(* IEC 61131-3 sources: plc-st-coding-agent/progress/evidence/f14_v5_public_pilot_20261112/jobs/codex_deepseek-v4pro, 18 files *)

(* ---- public-easy-01.candidate_01.st ---- *)
FUNCTION_BLOCK AutomatedFillingLineControl
VAR_INPUT
    bottleSensor : BOOL;
    cleaningConfirmButton : BOOL;
    fillingConfirmButton : BOOL;
    cappingConfirmButton : BOOL;
    packingConfirmButton : BOOL;
    finishedButton : BOOL;
END_VAR
VAR_OUTPUT
    Pump_Motor : BOOL;
    Filling_Valve : BOOL;
    Capping_Machine : BOOL;
    Packing_Machine : BOOL;
    Completion_Light : BOOL;
END_VAR
VAR
    State : INT := 0;
END_VAR

(* ENGINEERING_CONTRACT
- Pump_Motor: active from bottleSensor detection in Idle and latched through Cleaning; PUB003.
- Pump_Motor: deactivated when cleaningConfirmButton advances to Filling; PUB004.
- Filling_Valve: active from cleaningConfirmButton and held through Filling; PUB004.
- Filling_Valve: deactivated when fillingConfirmButton advances to Capping; PUB005.
- Capping_Machine: active from fillingConfirmButton and held through Capping; PUB005-PUB006.
- Capping_Machine: deactivated when cappingConfirmButton advances to Packing; PUB006.
- Packing_Machine: active from cappingConfirmButton and held through Packing; PUB006-PUB007.
- Packing_Machine: deactivated when packingConfirmButton lights Completion_Light; PUB007.
- Completion_Light: held until finishedButton resets it and returns to Idle; PUB007-PUB008.
- Level-checked inputs; only the current stage consumes its matching confirmation button.
- Same-scan priority: one stage transition per scan; output units are BOOL with no time bounds.
*)

CASE State OF
    0:
        Pump_Motor := FALSE;
        Filling_Valve := FALSE;
        Capping_Machine := FALSE;
        Packing_Machine := FALSE;
        Completion_Light := FALSE;

        IF bottleSensor THEN
            Pump_Motor := TRUE;
            State := 1;
        END_IF;

    1:
        Pump_Motor := TRUE;

        IF cleaningConfirmButton THEN
            Pump_Motor := FALSE;
            Filling_Valve := TRUE;
            State := 2;
        END_IF;

    2:
        Filling_Valve := TRUE;

        IF fillingConfirmButton THEN
            Filling_Valve := FALSE;
            Capping_Machine := TRUE;
            State := 3;
        END_IF;

    3:
        Capping_Machine := TRUE;

        IF cappingConfirmButton THEN
            Capping_Machine := FALSE;
            Packing_Machine := TRUE;
            State := 4;
        END_IF;

    4:
        Packing_Machine := TRUE;

        IF packingConfirmButton THEN
            Packing_Machine := FALSE;
            Completion_Light := TRUE;
            State := 5;
        END_IF;

    5:
        Completion_Light := TRUE;

        IF finishedButton THEN
            Completion_Light := FALSE;
            State := 0;
        END_IF;
END_CASE;

END_FUNCTION_BLOCK

(* ---- public-easy-01.candidate_02.st ---- *)
FUNCTION_BLOCK AutomatedFillingLineControl
VAR_INPUT
    bottleSensor : BOOL;
    cleaningConfirmButton : BOOL;
    fillingConfirmButton : BOOL;
    cappingConfirmButton : BOOL;
    packingConfirmButton : BOOL;
    finishedButton : BOOL;
END_VAR
VAR_OUTPUT
    Pump_Motor : BOOL;
    Filling_Valve : BOOL;
    Capping_Machine : BOOL;
    Packing_Machine : BOOL;
    Completion_Light : BOOL;
END_VAR
VAR
END_VAR

(* ENGINEERING_CONTRACT
- Pump_Motor: activated by bottleSensor, retained/holds until finishedButton reset; PUB003.
- Filling_Valve: activated by cleaningConfirmButton, retained until finishedButton reset; PUB004.
- Capping_Machine: activated by fillingConfirmButton, retained until finishedButton reset; PUB005.
- Packing_Machine: activated by cappingConfirmButton, retained until finishedButton reset; PUB006.
- Completion_Light: activated by packingConfirmButton, retained until finishedButton reset; PUB007.
- finishedButton: explicit common reset for all outputs, applied last in same scan; PUB008.
- Outputs are BOOL; no time bounds. Activation inputs are level-latched, not edge-only.
*)

IF bottleSensor THEN
    Pump_Motor := TRUE;
END_IF;

IF cleaningConfirmButton THEN
    Filling_Valve := TRUE;
END_IF;

IF fillingConfirmButton THEN
    Capping_Machine := TRUE;
END_IF;

IF cappingConfirmButton THEN
    Packing_Machine := TRUE;
END_IF;

IF packingConfirmButton THEN
    Completion_Light := TRUE;
END_IF;

IF finishedButton THEN
    Pump_Motor := FALSE;
    Filling_Valve := FALSE;
    Capping_Machine := FALSE;
    Packing_Machine := FALSE;
    Completion_Light := FALSE;
END_IF;

END_FUNCTION_BLOCK

(* ---- public-easy-01.raw_candidate_01.st ---- *)
FUNCTION_BLOCK AutomatedFillingLineControl
VAR_INPUT
    bottleSensor : BOOL;
    cleaningConfirmButton : BOOL;
    fillingConfirmButton : BOOL;
    cappingConfirmButton : BOOL;
    packingConfirmButton : BOOL;
    finishedButton : BOOL;
END_VAR
VAR_OUTPUT
    Pump_Motor : BOOL;
    Filling_Valve : BOOL;
    Capping_Machine : BOOL;
    Packing_Machine : BOOL;
    Completion_Light : BOOL;
END_VAR
VAR
    State : INT := 0;
END_VAR

(* ENGINEERING_CONTRACT
- Pump_Motor: active from bottleSensor detection in Idle and latched through Cleaning; PUB003.
- Pump_Motor: deactivated when cleaningConfirmButton advances to Filling; PUB004.
- Filling_Valve: active from cleaningConfirmButton and held through Filling; PUB004.
- Filling_Valve: deactivated when fillingConfirmButton advances to Capping; PUB005.
- Capping_Machine: active from fillingConfirmButton and held through Capping; PUB005-PUB006.
- Capping_Machine: deactivated when cappingConfirmButton advances to Packing; PUB006.
- Packing_Machine: active from cappingConfirmButton and held through Packing; PUB006-PUB007.
- Packing_Machine: deactivated when packingConfirmButton lights Completion_Light; PUB007.
- Completion_Light: held until finishedButton resets it and returns to Idle; PUB007-PUB008.
- Level-checked inputs; only the current stage consumes its matching confirmation button.
- Same-scan priority: one stage transition per scan; output units are BOOL with no time bounds.
*)

CASE State OF
    0:
        Pump_Motor := FALSE;
        Filling_Valve := FALSE;
        Capping_Machine := FALSE;
        Packing_Machine := FALSE;
        Completion_Light := FALSE;

        IF bottleSensor THEN
            Pump_Motor := TRUE;
            State := 1;
        END_IF;

    1:
        Pump_Motor := TRUE;

        IF cleaningConfirmButton THEN
            Pump_Motor := FALSE;
            Filling_Valve := TRUE;
            State := 2;
        END_IF;

    2:
        Filling_Valve := TRUE;

        IF fillingConfirmButton THEN
            Filling_Valve := FALSE;
            Capping_Machine := TRUE;
            State := 3;
        END_IF;

    3:
        Capping_Machine := TRUE;

        IF cappingConfirmButton THEN
            Capping_Machine := FALSE;
            Packing_Machine := TRUE;
            State := 4;
        END_IF;

    4:
        Packing_Machine := TRUE;

        IF packingConfirmButton THEN
            Packing_Machine := FALSE;
            Completion_Light := TRUE;
            State := 5;
        END_IF;

    5:
        Completion_Light := TRUE;

        IF finishedButton THEN
            Completion_Light := FALSE;
            State := 0;
        END_IF;
END_CASE;

END_FUNCTION_BLOCK

(* ---- public-easy-01.raw_candidate_02.st ---- *)
FUNCTION_BLOCK AutomatedFillingLineControl
VAR_INPUT
    bottleSensor : BOOL;
    cleaningConfirmButton : BOOL;
    fillingConfirmButton : BOOL;
    cappingConfirmButton : BOOL;
    packingConfirmButton : BOOL;
    finishedButton : BOOL;
END_VAR
VAR_OUTPUT
    Pump_Motor : BOOL;
    Filling_Valve : BOOL;
    Capping_Machine : BOOL;
    Packing_Machine : BOOL;
    Completion_Light : BOOL;
END_VAR
VAR
END_VAR

(* ENGINEERING_CONTRACT
- Pump_Motor: activated by bottleSensor, retained/holds until finishedButton reset; PUB003.
- Filling_Valve: activated by cleaningConfirmButton, retained until finishedButton reset; PUB004.
- Capping_Machine: activated by fillingConfirmButton, retained until finishedButton reset; PUB005.
- Packing_Machine: activated by cappingConfirmButton, retained until finishedButton reset; PUB006.
- Completion_Light: activated by packingConfirmButton, retained until finishedButton reset; PUB007.
- finishedButton: explicit common reset for all outputs, applied last in same scan; PUB008.
- Outputs are BOOL; no time bounds. Activation inputs are level-latched, not edge-only.
*)

IF bottleSensor THEN
    Pump_Motor := TRUE;
END_IF;

IF cleaningConfirmButton THEN
    Filling_Valve := TRUE;
END_IF;

IF fillingConfirmButton THEN
    Capping_Machine := TRUE;
END_IF;

IF cappingConfirmButton THEN
    Packing_Machine := TRUE;
END_IF;

IF packingConfirmButton THEN
    Completion_Light := TRUE;
END_IF;

IF finishedButton THEN
    Pump_Motor := FALSE;
    Filling_Valve := FALSE;
    Capping_Machine := FALSE;
    Packing_Machine := FALSE;
    Completion_Light := FALSE;
END_IF;

END_FUNCTION_BLOCK

(* ---- public-easy-04.candidate_01.st ---- *)
(*
ENGINEERING_CONTRACT
VFD_RUN [PUB002,PUB003,PUB006]: TRUE only while PASTE_E_STOP_NC=TRUE and the viscosity debounce timer has elapsed; same-scan emergency stop drops the run command and clears incomplete debounce timing; power-up state is OFF.
Debounce [PUB002,PUB003]: timer IN uses VISCOSITY_OK AND PASTE_E_STOP_NC with PT=DebounceTime; a FALSE viscosity input invalidates immediately, and a FALSE emergency stop resets incomplete timing.
Runtime [PUB004,PUB006]: adds TIME_TO_LTIME(CycleTime) once per invocation only while VFD_RUN=TRUE; preserves the accumulated value while stopped; starts at 0 ns.
Maintenance [PUB005,PUB006]: PUMP_MAINT_DUE becomes TRUE when accumulated runtime reaches 500 h; it is informational only, remains TRUE because runtime is monotonic, and does not affect run or safety logic; starts FALSE.
Units/boundaries: maintenance threshold uses T#500h with >= comparison; CycleTime and DebounceTime are assumed positive.
Unspecified: no reset is defined for accumulated runtime or the maintenance indication; non-positive input times follow normal TON/add behavior without additional clamping.
*)
FUNCTION_BLOCK JamPumpControl
VAR_INPUT
    VISCOSITY_OK : BOOL;
    PASTE_E_STOP_NC : BOOL;
    DebounceTime : TIME;
    CycleTime : TIME;
END_VAR
VAR_OUTPUT
    VFD_RUN : BOOL;
    PUMP_MAINT_DUE : BOOL;
    PUMP_RUNTIME_ACC : LTIME;
END_VAR
VAR
    tonViscosity : TON;
    RuntimeAcc : LTIME := LTIME#0s;
    MAINT_THRESHOLD : TIME := T#500h;
END_VAR

tonViscosity(IN := (VISCOSITY_OK AND PASTE_E_STOP_NC), PT := DebounceTime);

VFD_RUN := PASTE_E_STOP_NC AND tonViscosity.Q;

IF VFD_RUN THEN
    RuntimeAcc := RuntimeAcc + TIME_TO_LTIME(CycleTime);
END_IF;

PUMP_RUNTIME_ACC := RuntimeAcc;
PUMP_MAINT_DUE := PUMP_RUNTIME_ACC >= TIME_TO_LTIME(MAINT_THRESHOLD);

END_FUNCTION_BLOCK

(* ---- public-easy-04.raw_candidate_01.st ---- *)
(*
ENGINEERING_CONTRACT
VFD_RUN [PUB002,PUB003,PUB006]: TRUE only while PASTE_E_STOP_NC=TRUE and the viscosity debounce timer has elapsed; same-scan emergency stop drops the run command and clears incomplete debounce timing; power-up state is OFF.
Debounce [PUB002,PUB003]: timer IN uses VISCOSITY_OK AND PASTE_E_STOP_NC with PT=DebounceTime; a FALSE viscosity input invalidates immediately, and a FALSE emergency stop resets incomplete timing.
Runtime [PUB004,PUB006]: adds TIME_TO_LTIME(CycleTime) once per invocation only while VFD_RUN=TRUE; preserves the accumulated value while stopped; starts at 0 ns.
Maintenance [PUB005,PUB006]: PUMP_MAINT_DUE becomes TRUE when accumulated runtime reaches 500 h; it is informational only, remains TRUE because runtime is monotonic, and does not affect run or safety logic; starts FALSE.
Units/boundaries: maintenance threshold uses T#500h with >= comparison; CycleTime and DebounceTime are assumed positive.
Unspecified: no reset is defined for accumulated runtime or the maintenance indication; non-positive input times follow normal TON/add behavior without additional clamping.
*)
FUNCTION_BLOCK JamPumpControl
VAR_INPUT
    VISCOSITY_OK : BOOL;
    PASTE_E_STOP_NC : BOOL;
    DebounceTime : TIME;
    CycleTime : TIME;
END_VAR
VAR_OUTPUT
    VFD_RUN : BOOL;
    PUMP_MAINT_DUE : BOOL;
    PUMP_RUNTIME_ACC : LTIME;
END_VAR
VAR
    tonViscosity : TON;
    RuntimeAcc : LTIME := LTIME#0s;
    MAINT_THRESHOLD : TIME := T#500h;
END_VAR

tonViscosity(IN := (VISCOSITY_OK AND PASTE_E_STOP_NC), PT := DebounceTime);

VFD_RUN := PASTE_E_STOP_NC AND tonViscosity.Q;

IF VFD_RUN THEN
    RuntimeAcc := RuntimeAcc + TIME_TO_LTIME(CycleTime);
END_IF;

PUMP_RUNTIME_ACC := RuntimeAcc;
PUMP_MAINT_DUE := PUMP_RUNTIME_ACC >= TIME_TO_LTIME(MAINT_THRESHOLD);

END_FUNCTION_BLOCK

(* ---- public-hard-03.candidate_01.st ---- *)
TYPE ST_Recipe :
STRUCT
    recipeID : INT;
    ingredientType : INT;
    ingredientRatio : REAL;
    productionTemperature : REAL;
END_STRUCT
END_TYPE;

FUNCTION_BLOCK RecipeManagementSystem
(*
ENGINEERING_CONTRACT
- Operations are level-triggered; no edge or latch storage is added (PUB002-PUB006).
- recipeAdded/Deleted/Modified are active only during a successful selected scan; otherwise cleared.
- error/status clear each scan unless the selected operation reports a failure.
- Query retains the last successful recipeQueryResult; a missing recipe leaves it unchanged (PUB009).
- Add checks duplicate first, then smallest empty index, otherwise 16#8002/16#8003 (PUB010).
- Delete clears only recipeID in the matched slot (PUB011).
- Modify replaces the whole matched ST_Recipe with recipeIn (PUB012).
- recipeID=0 denotes an empty slot; searches ignore such slots (PUB008).
- Simultaneous requests use priority add > delete > modify > query (unspecified by task).
*)
VAR_INPUT
    addRecipe : BOOL;
    deleteRecipe : BOOL;
    modifyRecipe : BOOL;
    queryRecipe : BOOL;
    recipeIn : ST_Recipe;
END_VAR
VAR_OUTPUT
    recipeAdded : BOOL;
    recipeDeleted : BOOL;
    recipeModified : BOOL;
    recipeQueryResult : ST_Recipe;
    error : BOOL;
    status : WORD;
END_VAR
VAR_IN_OUT
    recipe : ARRAY[1..10] OF ST_Recipe;
END_VAR
VAR
    i : INT;
    foundIndex : INT;
    emptyIndex : INT;
    found : BOOL;
    emptyFound : BOOL;
END_VAR

recipeAdded := FALSE;
recipeDeleted := FALSE;
recipeModified := FALSE;
error := FALSE;
status := 0;

IF addRecipe THEN
    found := FALSE;
    foundIndex := 0;
    FOR i := 1 TO 10 DO
        IF (recipe[i].recipeID <> 0) AND (recipe[i].recipeID = recipeIn.recipeID) THEN
            found := TRUE;
            foundIndex := i;
            EXIT;
        END_IF;
    END_FOR;

    IF found THEN
        error := TRUE;
        status := WORD#16#8002;
    ELSE
        emptyFound := FALSE;
        emptyIndex := 0;
        FOR i := 1 TO 10 DO
            IF recipe[i].recipeID = 0 THEN
                emptyFound := TRUE;
                emptyIndex := i;
                EXIT;
            END_IF;
        END_FOR;

        IF NOT emptyFound THEN
            error := TRUE;
            status := WORD#16#8003;
        ELSE
            recipe[emptyIndex].recipeID := recipeIn.recipeID;
            recipe[emptyIndex].ingredientType := recipeIn.ingredientType;
            recipe[emptyIndex].ingredientRatio := recipeIn.ingredientRatio;
            recipe[emptyIndex].productionTemperature := recipeIn.productionTemperature;
            recipeAdded := TRUE;
            error := FALSE;
            status := 0;
        END_IF;
    END_IF;

ELSIF deleteRecipe THEN
    found := FALSE;
    foundIndex := 0;
    FOR i := 1 TO 10 DO
        IF (recipe[i].recipeID <> 0) AND (recipe[i].recipeID = recipeIn.recipeID) THEN
            found := TRUE;
            foundIndex := i;
            EXIT;
        END_IF;
    END_FOR;

    IF NOT found THEN
        error := TRUE;
        status := WORD#16#8004;
    ELSE
        recipe[foundIndex].recipeID := 0;
        recipeDeleted := TRUE;
        error := FALSE;
        status := 0;
    END_IF;

ELSIF modifyRecipe THEN
    found := FALSE;
    foundIndex := 0;
    FOR i := 1 TO 10 DO
        IF (recipe[i].recipeID <> 0) AND (recipe[i].recipeID = recipeIn.recipeID) THEN
            found := TRUE;
            foundIndex := i;
            EXIT;
        END_IF;
    END_FOR;

    IF NOT found THEN
        error := TRUE;
        status := WORD#16#8005;
    ELSE
        recipe[foundIndex] := recipeIn;
        recipeModified := TRUE;
        error := FALSE;
        status := 0;
    END_IF;

ELSIF queryRecipe THEN
    found := FALSE;
    foundIndex := 0;
    FOR i := 1 TO 10 DO
        IF (recipe[i].recipeID <> 0) AND (recipe[i].recipeID = recipeIn.recipeID) THEN
            found := TRUE;
            foundIndex := i;
            EXIT;
        END_IF;
    END_FOR;

    IF NOT found THEN
        error := TRUE;
        status := WORD#16#8001;
    ELSE
        recipeQueryResult := recipe[foundIndex];
        error := FALSE;
        status := 0;
    END_IF;
END_IF;

END_FUNCTION_BLOCK

(* ---- public-hard-03.candidate_02.st ---- *)
TYPE ST_Recipe :
STRUCT
    recipeID : INT;
    ingredientType : INT;
    ingredientRatio : REAL;
    productionTemperature : REAL;
END_STRUCT
END_TYPE;

FUNCTION_BLOCK RecipeManagementSystem
(*
ENGINEERING_CONTRACT
- Request inputs are level-triggered; no edge or latch storage is added.
- recipeAdded/recipeDeleted/recipeModified are true only on a successful scan of the matching request, otherwise false.
- error/status clear at scan start; any failed request in the scan sets them.
- Query success overwrites recipeQueryResult; a failed query leaves it unchanged.
- Add checks duplicate first, then finds the smallest empty index, then checks full database.
- Delete clears only recipeID in the matched slot.
- Modify replaces the entire matched ST_Recipe with recipeIn.
- Empty slots are identified by recipeID = 0 and are ignored during normal searches.
- Simultaneous requests are unspecified; they are evaluated in interface order add/delete/modify/query.
*)
VAR_INPUT
    addRecipe : BOOL;
    deleteRecipe : BOOL;
    modifyRecipe : BOOL;
    queryRecipe : BOOL;
    recipeIn : ST_Recipe;
END_VAR
VAR_OUTPUT
    recipeAdded : BOOL;
    recipeDeleted : BOOL;
    recipeModified : BOOL;
    recipeQueryResult : ST_Recipe;
    error : BOOL;
    status : WORD;
END_VAR
VAR_IN_OUT
    recipe : ARRAY[1..10] OF ST_Recipe;
END_VAR
VAR
    i : INT;
    foundIndex : INT;
    emptyIndex : INT;
    found : BOOL;
    emptyFound : BOOL;
END_VAR

recipeAdded := FALSE;
recipeDeleted := FALSE;
recipeModified := FALSE;
error := FALSE;
status := 0;

IF addRecipe THEN
    found := FALSE;
    foundIndex := 0;
    FOR i := 1 TO 10 DO
        IF (recipe[i].recipeID <> 0) AND (recipe[i].recipeID = recipeIn.recipeID) THEN
            found := TRUE;
            foundIndex := i;
            EXIT;
        END_IF;
    END_FOR;

    IF found THEN
        error := TRUE;
        status := WORD#16#8002;
    ELSE
        emptyFound := FALSE;
        emptyIndex := 0;
        FOR i := 1 TO 10 DO
            IF recipe[i].recipeID = 0 THEN
                emptyFound := TRUE;
                emptyIndex := i;
                EXIT;
            END_IF;
        END_FOR;

        IF NOT emptyFound THEN
            error := TRUE;
            status := WORD#16#8003;
        ELSE
            recipe[emptyIndex].recipeID := recipeIn.recipeID;
            recipe[emptyIndex].ingredientType := recipeIn.ingredientType;
            recipe[emptyIndex].ingredientRatio := recipeIn.ingredientRatio;
            recipe[emptyIndex].productionTemperature := recipeIn.productionTemperature;
            recipeAdded := TRUE;
        END_IF;
    END_IF;
END_IF;

IF deleteRecipe THEN
    found := FALSE;
    foundIndex := 0;
    FOR i := 1 TO 10 DO
        IF (recipe[i].recipeID <> 0) AND (recipe[i].recipeID = recipeIn.recipeID) THEN
            found := TRUE;
            foundIndex := i;
            EXIT;
        END_IF;
    END_FOR;

    IF NOT found THEN
        error := TRUE;
        status := WORD#16#8004;
    ELSE
        recipe[foundIndex].recipeID := 0;
        recipeDeleted := TRUE;
    END_IF;
END_IF;

IF modifyRecipe THEN
    found := FALSE;
    foundIndex := 0;
    FOR i := 1 TO 10 DO
        IF (recipe[i].recipeID <> 0) AND (recipe[i].recipeID = recipeIn.recipeID) THEN
            found := TRUE;
            foundIndex := i;
            EXIT;
        END_IF;
    END_FOR;

    IF NOT found THEN
        error := TRUE;
        status := WORD#16#8005;
    ELSE
        recipe[foundIndex] := recipeIn;
        recipeModified := TRUE;
    END_IF;
END_IF;

IF queryRecipe THEN
    found := FALSE;
    foundIndex := 0;
    FOR i := 1 TO 10 DO
        IF (recipe[i].recipeID <> 0) AND (recipe[i].recipeID = recipeIn.recipeID) THEN
            found := TRUE;
            foundIndex := i;
            EXIT;
        END_IF;
    END_FOR;

    IF NOT found THEN
        error := TRUE;
        status := WORD#16#8001;
    ELSE
        recipeQueryResult := recipe[foundIndex];
    END_IF;
END_IF;

END_FUNCTION_BLOCK

(* ---- public-hard-03.raw_candidate_01.st ---- *)
TYPE ST_Recipe :
STRUCT
    recipeID : INT;
    ingredientType : INT;
    ingredientRatio : REAL;
    productionTemperature : REAL;
END_STRUCT
END_TYPE

FUNCTION_BLOCK RecipeManagementSystem
(*
ENGINEERING_CONTRACT
- Operations are level-triggered; no edge or latch storage is added (PUB002-PUB006).
- recipeAdded/Deleted/Modified are active only during a successful selected scan; otherwise cleared.
- error/status clear each scan unless the selected operation reports a failure.
- Query retains the last successful recipeQueryResult; a missing recipe leaves it unchanged (PUB009).
- Add checks duplicate first, then smallest empty index, otherwise 16#8002/16#8003 (PUB010).
- Delete clears only recipeID in the matched slot (PUB011).
- Modify replaces the whole matched ST_Recipe with recipeIn (PUB012).
- recipeID=0 denotes an empty slot; searches ignore such slots (PUB008).
- Simultaneous requests use priority add > delete > modify > query (unspecified by task).
*)
VAR_INPUT
    addRecipe : BOOL;
    deleteRecipe : BOOL;
    modifyRecipe : BOOL;
    queryRecipe : BOOL;
    recipeIn : ST_Recipe;
END_VAR
VAR_OUTPUT
    recipeAdded : BOOL;
    recipeDeleted : BOOL;
    recipeModified : BOOL;
    recipeQueryResult : ST_Recipe;
    error : BOOL;
    status : WORD;
END_VAR
VAR_IN_OUT
    recipe : ARRAY[1..10] OF ST_Recipe;
END_VAR
VAR
    i : INT;
    foundIndex : INT;
    emptyIndex : INT;
    found : BOOL;
    emptyFound : BOOL;
END_VAR

recipeAdded := FALSE;
recipeDeleted := FALSE;
recipeModified := FALSE;
error := FALSE;
status := 0;

IF addRecipe THEN
    found := FALSE;
    foundIndex := 0;
    FOR i := 1 TO 10 DO
        IF (recipe[i].recipeID <> 0) AND (recipe[i].recipeID = recipeIn.recipeID) THEN
            found := TRUE;
            foundIndex := i;
            EXIT;
        END_IF;
    END_FOR;

    IF found THEN
        error := TRUE;
        status := WORD#16#8002;
    ELSE
        emptyFound := FALSE;
        emptyIndex := 0;
        FOR i := 1 TO 10 DO
            IF recipe[i].recipeID = 0 THEN
                emptyFound := TRUE;
                emptyIndex := i;
                EXIT;
            END_IF;
        END_FOR;

        IF NOT emptyFound THEN
            error := TRUE;
            status := WORD#16#8003;
        ELSE
            recipe[emptyIndex].recipeID := recipeIn.recipeID;
            recipe[emptyIndex].ingredientType := recipeIn.ingredientType;
            recipe[emptyIndex].ingredientRatio := recipeIn.ingredientRatio;
            recipe[emptyIndex].productionTemperature := recipeIn.productionTemperature;
            recipeAdded := TRUE;
            error := FALSE;
            status := 0;
        END_IF;
    END_IF;

ELSIF deleteRecipe THEN
    found := FALSE;
    foundIndex := 0;
    FOR i := 1 TO 10 DO
        IF (recipe[i].recipeID <> 0) AND (recipe[i].recipeID = recipeIn.recipeID) THEN
            found := TRUE;
            foundIndex := i;
            EXIT;
        END_IF;
    END_FOR;

    IF NOT found THEN
        error := TRUE;
        status := WORD#16#8004;
    ELSE
        recipe[foundIndex].recipeID := 0;
        recipeDeleted := TRUE;
        error := FALSE;
        status := 0;
    END_IF;

ELSIF modifyRecipe THEN
    found := FALSE;
    foundIndex := 0;
    FOR i := 1 TO 10 DO
        IF (recipe[i].recipeID <> 0) AND (recipe[i].recipeID = recipeIn.recipeID) THEN
            found := TRUE;
            foundIndex := i;
            EXIT;
        END_IF;
    END_FOR;

    IF NOT found THEN
        error := TRUE;
        status := WORD#16#8005;
    ELSE
        recipe[foundIndex] := recipeIn;
        recipeModified := TRUE;
        error := FALSE;
        status := 0;
    END_IF;

ELSIF queryRecipe THEN
    found := FALSE;
    foundIndex := 0;
    FOR i := 1 TO 10 DO
        IF (recipe[i].recipeID <> 0) AND (recipe[i].recipeID = recipeIn.recipeID) THEN
            found := TRUE;
            foundIndex := i;
            EXIT;
        END_IF;
    END_FOR;

    IF NOT found THEN
        error := TRUE;
        status := WORD#16#8001;
    ELSE
        recipeQueryResult := recipe[foundIndex];
        error := FALSE;
        status := 0;
    END_IF;
END_IF;

END_FUNCTION_BLOCK

(* ---- public-hard-03.raw_candidate_02.st ---- *)
TYPE ST_Recipe :
STRUCT
    recipeID : INT;
    ingredientType : INT;
    ingredientRatio : REAL;
    productionTemperature : REAL;
END_STRUCT
END_TYPE;

FUNCTION_BLOCK RecipeManagementSystem
(*
ENGINEERING_CONTRACT
- Request inputs are level-triggered; no edge or latch storage is added.
- recipeAdded/recipeDeleted/recipeModified are true only on a successful scan of the matching request, otherwise false.
- error/status clear at scan start; any failed request in the scan sets them.
- Query success overwrites recipeQueryResult; a failed query leaves it unchanged.
- Add checks duplicate first, then finds the smallest empty index, then checks full database.
- Delete clears only recipeID in the matched slot.
- Modify replaces the entire matched ST_Recipe with recipeIn.
- Empty slots are identified by recipeID = 0 and are ignored during normal searches.
- Simultaneous requests are unspecified; they are evaluated in interface order add/delete/modify/query.
*)
VAR_INPUT
    addRecipe : BOOL;
    deleteRecipe : BOOL;
    modifyRecipe : BOOL;
    queryRecipe : BOOL;
    recipeIn : ST_Recipe;
END_VAR
VAR_OUTPUT
    recipeAdded : BOOL;
    recipeDeleted : BOOL;
    recipeModified : BOOL;
    recipeQueryResult : ST_Recipe;
    error : BOOL;
    status : WORD;
END_VAR
VAR_IN_OUT
    recipe : ARRAY[1..10] OF ST_Recipe;
END_VAR
VAR
    i : INT;
    foundIndex : INT;
    emptyIndex : INT;
    found : BOOL;
    emptyFound : BOOL;
END_VAR

recipeAdded := FALSE;
recipeDeleted := FALSE;
recipeModified := FALSE;
error := FALSE;
status := 0;

IF addRecipe THEN
    found := FALSE;
    foundIndex := 0;
    FOR i := 1 TO 10 DO
        IF (recipe[i].recipeID <> 0) AND (recipe[i].recipeID = recipeIn.recipeID) THEN
            found := TRUE;
            foundIndex := i;
            EXIT;
        END_IF;
    END_FOR;

    IF found THEN
        error := TRUE;
        status := WORD#16#8002;
    ELSE
        emptyFound := FALSE;
        emptyIndex := 0;
        FOR i := 1 TO 10 DO
            IF recipe[i].recipeID = 0 THEN
                emptyFound := TRUE;
                emptyIndex := i;
                EXIT;
            END_IF;
        END_FOR;

        IF NOT emptyFound THEN
            error := TRUE;
            status := WORD#16#8003;
        ELSE
            recipe[emptyIndex].recipeID := recipeIn.recipeID;
            recipe[emptyIndex].ingredientType := recipeIn.ingredientType;
            recipe[emptyIndex].ingredientRatio := recipeIn.ingredientRatio;
            recipe[emptyIndex].productionTemperature := recipeIn.productionTemperature;
            recipeAdded := TRUE;
        END_IF;
    END_IF;
END_IF;

IF deleteRecipe THEN
    found := FALSE;
    foundIndex := 0;
    FOR i := 1 TO 10 DO
        IF (recipe[i].recipeID <> 0) AND (recipe[i].recipeID = recipeIn.recipeID) THEN
            found := TRUE;
            foundIndex := i;
            EXIT;
        END_IF;
    END_FOR;

    IF NOT found THEN
        error := TRUE;
        status := WORD#16#8004;
    ELSE
        recipe[foundIndex].recipeID := 0;
        recipeDeleted := TRUE;
    END_IF;
END_IF;

IF modifyRecipe THEN
    found := FALSE;
    foundIndex := 0;
    FOR i := 1 TO 10 DO
        IF (recipe[i].recipeID <> 0) AND (recipe[i].recipeID = recipeIn.recipeID) THEN
            found := TRUE;
            foundIndex := i;
            EXIT;
        END_IF;
    END_FOR;

    IF NOT found THEN
        error := TRUE;
        status := WORD#16#8005;
    ELSE
        recipe[foundIndex] := recipeIn;
        recipeModified := TRUE;
    END_IF;
END_IF;

IF queryRecipe THEN
    found := FALSE;
    foundIndex := 0;
    FOR i := 1 TO 10 DO
        IF (recipe[i].recipeID <> 0) AND (recipe[i].recipeID = recipeIn.recipeID) THEN
            found := TRUE;
            foundIndex := i;
            EXIT;
        END_IF;
    END_FOR;

    IF NOT found THEN
        error := TRUE;
        status := WORD#16#8001;
    ELSE
        recipeQueryResult := recipe[foundIndex];
    END_IF;
END_IF;

END_FUNCTION_BLOCK

(* ---- public-medium-03.candidate_01.st ---- *)
(* ENGINEERING_CONTRACT
   average: recomputed each scan for active stored samples; 0.0 when no samples or after reset. Units follow value.
   windowSizeReached: TRUE iff stored valid sample count >= current valid windowSize; cleared by reset and on invalid window.
   error/status: enabled by windowSize outside 1..100; status 16#8200, otherwise 16#0000 (PUB004/PUB006/PUB007).
   same-scan priority: level-true reset first, then window validation, then cyclic or rising-edge sample; cyclic TRUE ignores trigger edge (PUB002/PUB003).
   reset: explicit level-true clear of stored samples, count, average, and reached state; no same-scan sample after reset.
   trigger: internal rising-edge detector; each valid, non-reset rising edge adds one value.
   retention: valid stored samples persist without reset; dynamic window resizing uses the newest min(validCount, windowSize) samples.
   boundaries: windowSize [1,100], storage capacity 100; average is LREAL mean with no unit conversion.
*)
FUNCTION_BLOCK FB
VAR_INPUT
    cyclicExecution : BOOL;
    trigger : BOOL;
    value : LREAL;
    windowSize : INT;
    reset : BOOL;
END_VAR
VAR_OUTPUT
    average : LREAL;
    windowSizeReached : BOOL;
    error : BOOL;
    status : WORD;
END_VAR
VAR
    buffer : ARRAY[0..99] OF LREAL;
    nextIndex : INT := 0;
    validCount : INT := 0;
    triggerPrevious : BOOL;
    triggerRising : BOOL;
    activeWindow : INT;
    startIndex : INT;
    loopIndex : INT;
    sumValue : LREAL;
END_VAR

triggerRising := trigger AND NOT triggerPrevious;
triggerPrevious := trigger;

IF reset THEN
    validCount := 0;
    nextIndex := 0;
    average := 0.0;
    windowSizeReached := FALSE;
END_IF;

IF (windowSize < 1) OR (windowSize > 100) THEN
    error := TRUE;
    status := 16#8200;
    average := 0.0;
    windowSizeReached := FALSE;
ELSE
    error := FALSE;
    status := 16#0000;

    IF NOT reset THEN
        IF cyclicExecution OR triggerRising THEN
            buffer[nextIndex] := value;
            nextIndex := nextIndex + 1;

            IF nextIndex > 99 THEN
                nextIndex := 0;
            END_IF;

            IF validCount < 100 THEN
                validCount := validCount + 1;
            END_IF;
        END_IF;
    END_IF;

    activeWindow := windowSize;
    IF activeWindow > validCount THEN
        activeWindow := validCount;
    END_IF;

    IF activeWindow > 0 THEN
        sumValue := 0.0;
        FOR loopIndex := 0 TO activeWindow - 1 DO
            startIndex := nextIndex - 1 - loopIndex;
            IF startIndex < 0 THEN
                startIndex := startIndex + 100;
            END_IF;
            sumValue := sumValue + buffer[startIndex];
        END_FOR;
        average := sumValue / INT_TO_LREAL(activeWindow);
    ELSE
        average := 0.0;
    END_IF;

    windowSizeReached := validCount >= windowSize;
END_IF;
END_FUNCTION_BLOCK

(* ---- public-medium-03.raw_candidate_01.st ---- *)
(* ENGINEERING_CONTRACT
   average: recomputed each scan for active stored samples; 0.0 when no samples or after reset. Units follow value.
   windowSizeReached: TRUE iff stored valid sample count >= current valid windowSize; cleared by reset and on invalid window.
   error/status: enabled by windowSize outside 1..100; status 16#8200, otherwise 16#0000 (PUB004/PUB006/PUB007).
   same-scan priority: level-true reset first, then window validation, then cyclic or rising-edge sample; cyclic TRUE ignores trigger edge (PUB002/PUB003).
   reset: explicit level-true clear of stored samples, count, average, and reached state; no same-scan sample after reset.
   trigger: internal rising-edge detector; each valid, non-reset rising edge adds one value.
   retention: valid stored samples persist without reset; dynamic window resizing uses the newest min(validCount, windowSize) samples.
   boundaries: windowSize [1,100], storage capacity 100; average is LREAL mean with no unit conversion.
*)
FUNCTION_BLOCK FB
VAR_INPUT
    cyclicExecution : BOOL;
    trigger : BOOL;
    value : LREAL;
    windowSize : INT;
    reset : BOOL;
END_VAR
VAR_OUTPUT
    average : LREAL;
    windowSizeReached : BOOL;
    error : BOOL;
    status : WORD;
END_VAR
VAR
    buffer : ARRAY[0..99] OF LREAL;
    nextIndex : INT := 0;
    validCount : INT := 0;
    triggerPrevious : BOOL;
    triggerRising : BOOL;
    activeWindow : INT;
    startIndex : INT;
    loopIndex : INT;
    sumValue : LREAL;
END_VAR

triggerRising := trigger AND NOT triggerPrevious;
triggerPrevious := trigger;

IF reset THEN
    validCount := 0;
    nextIndex := 0;
    average := 0.0;
    windowSizeReached := FALSE;
END_IF;

IF (windowSize < 1) OR (windowSize > 100) THEN
    error := TRUE;
    status := 16#8200;
    average := 0.0;
    windowSizeReached := FALSE;
ELSE
    error := FALSE;
    status := 16#0000;

    IF NOT reset THEN
        IF cyclicExecution OR triggerRising THEN
            buffer[nextIndex] := value;
            nextIndex := nextIndex + 1;

            IF nextIndex > 99 THEN
                nextIndex := 0;
            END_IF;

            IF validCount < 100 THEN
                validCount := validCount + 1;
            END_IF;
        END_IF;
    END_IF;

    activeWindow := windowSize;
    IF activeWindow > validCount THEN
        activeWindow := validCount;
    END_IF;

    IF activeWindow > 0 THEN
        sumValue := 0.0;
        FOR loopIndex := 0 TO activeWindow - 1 DO
            startIndex := nextIndex - 1 - loopIndex;
            IF startIndex < 0 THEN
                startIndex := startIndex + 100;
            END_IF;
            sumValue := sumValue + buffer[startIndex];
        END_FOR;
        average := sumValue / INT_TO_LREAL(activeWindow);
    ELSE
        average := 0.0;
    END_IF;

    windowSizeReached := validCount >= windowSize;
END_IF;
END_FUNCTION_BLOCK

(* ---- public-medium-04.candidate_01.st ---- *)
FUNCTION_BLOCK FB_TemperatureControl
VAR_INPUT
    TemperatureSensorInput : REAL;
    SetTemperature : REAL;
END_VAR
VAR_OUTPUT
    CurrentTemperature : REAL;
    SetTempDisplay : REAL;
    HeaterStatus : BOOL;
    OverheatProtection : BOOL;
    HeaterOutput : BOOL;
END_VAR
VAR
    SensorFault : BOOL;
    HeatRunTimer : TON;
    CoolDownTimer : TON;
END_VAR

(* ENGINEERING_CONTRACT
- CurrentTemperature/SetTempDisplay: copied from inputs every scan (PUB001, PUB002, PUB007); no retention; REAL.
- HeaterStatus: ON only while HeaterOutput is ON; no latch; cleared with heater OFF, overheat, or fault; same-scan as HeaterOutput; BOOL.
- OverheatProtection: latched when continuous heater run reaches >= T#5S (PUB006); held during T#3S cooldown; auto-clears after cooldown; BOOL.
- HeaterOutput: ON when no fault and actual < set (PUB003, PUB004); OFF when actual >= set, sensor fault, or protection (PUB005, PUB007, PUB008).
- SensorFault: TRUE when input < 0.0 or > 100.0 (PUB008); forces heater OFF; does not reset an active overheat cooldown.
- Unspecified: actual = set is interpreted as OFF; no hysteresis; after T#3S cooldown, normal control resumes automatically.
*)

CurrentTemperature := TemperatureSensorInput;
SetTempDisplay := SetTemperature;

SensorFault := (TemperatureSensorInput < 0.0) OR (TemperatureSensorInput > 100.0);

IF SensorFault THEN
    HeaterOutput := FALSE;
    HeaterStatus := FALSE;
    HeatRunTimer(IN := FALSE, PT := T#5S);

    IF OverheatProtection THEN
        CoolDownTimer(IN := TRUE, PT := T#3S);
        IF CoolDownTimer.Q THEN
            OverheatProtection := FALSE;
        END_IF;
    ELSE
        CoolDownTimer(IN := FALSE, PT := T#3S);
    END_IF;

ELSE
    IF OverheatProtection THEN
        HeaterOutput := FALSE;
        HeaterStatus := FALSE;
        HeatRunTimer(IN := FALSE, PT := T#5S);
        CoolDownTimer(IN := TRUE, PT := T#3S);

        IF CoolDownTimer.Q THEN
            OverheatProtection := FALSE;
        END_IF;

    ELSE
        IF TemperatureSensorInput < SetTemperature THEN
            HeaterOutput := TRUE;
            HeaterStatus := TRUE;
            HeatRunTimer(IN := TRUE, PT := T#5S);
            CoolDownTimer(IN := FALSE, PT := T#3S);

            IF HeatRunTimer.Q THEN
                OverheatProtection := TRUE;
                HeaterOutput := FALSE;
                HeaterStatus := FALSE;
            END_IF;

        ELSE
            HeaterOutput := FALSE;
            HeaterStatus := FALSE;
            HeatRunTimer(IN := FALSE, PT := T#5S);
            CoolDownTimer(IN := FALSE, PT := T#3S);
        END_IF;
    END_IF;
END_IF;

END_FUNCTION_BLOCK

(* ---- public-medium-04.candidate_02.st ---- *)
FUNCTION_BLOCK FB_TemperatureControl
VAR_INPUT
    TemperatureSensorInput : REAL;
    SetTemperature : REAL;
END_VAR
VAR_OUTPUT
    CurrentTemperature : REAL;
    SetTempDisplay : REAL;
    HeaterStatus : BOOL;
    OverheatProtection : BOOL;
    HeaterOutput : BOOL;
END_VAR
VAR
    SensorFault : BOOL;
    FreeClock : TON;
    HeatStartTime : TIME;
    HeatWasRunning : BOOL;
    HeatElapsed : TIME;
    CooldownStartTime : TIME;
    CoolElapsed : TIME;
END_VAR

(* ENGINEERING_CONTRACT
- CurrentTemperature/SetTempDisplay: copied from inputs every scan (PUB001, PUB002, PUB007); REAL.
- SensorFault: TRUE only when input < 0.0 or > 100.0 (PUB008); forces heater off.
- HeaterOutput/HeaterStatus: ON when no fault, no overheat, and actual < set; OFF at actual >= set (PUB003-PUB005, PUB007).
- OverheatProtection: latched after continuous heat > T#5S; held during cooldown; cleared when cooldown >= T#3S, then normal control is evaluated same scan (PUB006).
- Cooldown continues during sensor fault; heater remains off while fault is active.
- Timing: free-running TIME clock with snapshots; strict > for overheat, >= for cooldown clearance.
*)

CurrentTemperature := TemperatureSensorInput;
SetTempDisplay := SetTemperature;

SensorFault := (TemperatureSensorInput < 0.0) OR (TemperatureSensorInput > 100.0);

FreeClock(IN := TRUE, PT := T#60M);

IF OverheatProtection THEN
    CoolElapsed := FreeClock.ET - CooldownStartTime;
    IF CoolElapsed >= T#3S THEN
        OverheatProtection := FALSE;
    END_IF;
END_IF;

IF SensorFault OR OverheatProtection THEN
    HeaterOutput := FALSE;
    HeatWasRunning := FALSE;
ELSIF TemperatureSensorInput < SetTemperature THEN
    IF NOT HeatWasRunning THEN
        HeatStartTime := FreeClock.ET;
        HeatWasRunning := TRUE;
    END_IF;

    HeatElapsed := FreeClock.ET - HeatStartTime;

    IF HeatElapsed > T#5S THEN
        OverheatProtection := TRUE;
        CooldownStartTime := FreeClock.ET;
        HeatWasRunning := FALSE;
        HeaterOutput := FALSE;
    ELSE
        HeaterOutput := TRUE;
    END_IF;
ELSE
    HeatWasRunning := FALSE;
    HeaterOutput := FALSE;
END_IF;

HeaterStatus := HeaterOutput;

END_FUNCTION_BLOCK

(* ---- public-medium-04.raw_candidate_01.st ---- *)
FUNCTION_BLOCK FB_TemperatureControl
VAR_INPUT
    TemperatureSensorInput : REAL;
    SetTemperature : REAL;
END_VAR
VAR_OUTPUT
    CurrentTemperature : REAL;
    SetTempDisplay : REAL;
    HeaterStatus : BOOL;
    OverheatProtection : BOOL;
    HeaterOutput : BOOL;
END_VAR
VAR
    SensorFault : BOOL;
    HeatRunTimer : TON;
    CoolDownTimer : TON;
END_VAR

(* ENGINEERING_CONTRACT
- CurrentTemperature/SetTempDisplay: copied from inputs every scan (PUB001, PUB002, PUB007); no retention; REAL.
- HeaterStatus: ON only while HeaterOutput is ON; no latch; cleared with heater OFF, overheat, or fault; same-scan as HeaterOutput; BOOL.
- OverheatProtection: latched when continuous heater run reaches >= T#5S (PUB006); held during T#3S cooldown; auto-clears after cooldown; BOOL.
- HeaterOutput: ON when no fault and actual < set (PUB003, PUB004); OFF when actual >= set, sensor fault, or protection (PUB005, PUB007, PUB008).
- SensorFault: TRUE when input < 0.0 or > 100.0 (PUB008); forces heater OFF; does not reset an active overheat cooldown.
- Unspecified: actual = set is interpreted as OFF; no hysteresis; after T#3S cooldown, normal control resumes automatically.
*)

CurrentTemperature := TemperatureSensorInput;
SetTempDisplay := SetTemperature;

SensorFault := (TemperatureSensorInput < 0.0) OR (TemperatureSensorInput > 100.0);

IF SensorFault THEN
    HeaterOutput := FALSE;
    HeaterStatus := FALSE;
    HeatRunTimer(IN := FALSE, PT := T#5S);

    IF OverheatProtection THEN
        CoolDownTimer(IN := TRUE, PT := T#3S);
        IF CoolDownTimer.Q THEN
            OverheatProtection := FALSE;
        END_IF
    ELSE
        CoolDownTimer(IN := FALSE, PT := T#3S);
    END_IF

ELSE
    IF OverheatProtection THEN
        HeaterOutput := FALSE;
        HeaterStatus := FALSE;
        HeatRunTimer(IN := FALSE, PT := T#5S);
        CoolDownTimer(IN := TRUE, PT := T#3S);

        IF CoolDownTimer.Q THEN
            OverheatProtection := FALSE;
        END_IF

    ELSE
        IF TemperatureSensorInput < SetTemperature THEN
            HeaterOutput := TRUE;
            HeaterStatus := TRUE;
            HeatRunTimer(IN := TRUE, PT := T#5S);
            CoolDownTimer(IN := FALSE, PT := T#3S);

            IF HeatRunTimer.Q THEN
                OverheatProtection := TRUE;
                HeaterOutput := FALSE;
                HeaterStatus := FALSE;
            END_IF

        ELSE
            HeaterOutput := FALSE;
            HeaterStatus := FALSE;
            HeatRunTimer(IN := FALSE, PT := T#5S);
            CoolDownTimer(IN := FALSE, PT := T#3S);
        END_IF
    END_IF
END_IF

END_FUNCTION_BLOCK

(* ---- public-medium-04.raw_candidate_02.st ---- *)
FUNCTION_BLOCK FB_TemperatureControl
VAR_INPUT
    TemperatureSensorInput : REAL;
    SetTemperature : REAL;
END_VAR
VAR_OUTPUT
    CurrentTemperature : REAL;
    SetTempDisplay : REAL;
    HeaterStatus : BOOL;
    OverheatProtection : BOOL;
    HeaterOutput : BOOL;
END_VAR
VAR
    SensorFault : BOOL;
    FreeClock : TON;
    HeatStartTime : TIME;
    HeatWasRunning : BOOL;
    HeatElapsed : TIME;
    CooldownStartTime : TIME;
    CoolElapsed : TIME;
END_VAR

(* ENGINEERING_CONTRACT
- CurrentTemperature/SetTempDisplay: copied from inputs every scan (PUB001, PUB002, PUB007); REAL.
- SensorFault: TRUE only when input < 0.0 or > 100.0 (PUB008); forces heater off.
- HeaterOutput/HeaterStatus: ON when no fault, no overheat, and actual < set; OFF at actual >= set (PUB003-PUB005, PUB007).
- OverheatProtection: latched after continuous heat > T#5S; held during cooldown; cleared when cooldown >= T#3S, then normal control is evaluated same scan (PUB006).
- Cooldown continues during sensor fault; heater remains off while fault is active.
- Timing: free-running TIME clock with snapshots; strict > for overheat, >= for cooldown clearance.
*)

CurrentTemperature := TemperatureSensorInput;
SetTempDisplay := SetTemperature;

SensorFault := (TemperatureSensorInput < 0.0) OR (TemperatureSensorInput > 100.0);

FreeClock(IN := TRUE, PT := T#60M);

IF OverheatProtection THEN
    CoolElapsed := FreeClock.ET - CooldownStartTime;
    IF CoolElapsed >= T#3S THEN
        OverheatProtection := FALSE;
    END_IF;
END_IF;

IF SensorFault OR OverheatProtection THEN
    HeaterOutput := FALSE;
    HeatWasRunning := FALSE;
ELSIF TemperatureSensorInput < SetTemperature THEN
    IF NOT HeatWasRunning THEN
        HeatStartTime := FreeClock.ET;
        HeatWasRunning := TRUE;
    END_IF;

    HeatElapsed := FreeClock.ET - HeatStartTime;

    IF HeatElapsed > T#5S THEN
        OverheatProtection := TRUE;
        CooldownStartTime := FreeClock.ET;
        HeatWasRunning := FALSE;
        HeaterOutput := FALSE;
    ELSE
        HeaterOutput := TRUE;
    END_IF;
ELSE
    HeatWasRunning := FALSE;
    HeaterOutput := FALSE;
END_IF;

HeaterStatus := HeaterOutput;

END_FUNCTION_BLOCK

(* ---- public-medium-08.candidate_01.st ---- *)
(* ENGINEERING_CONTRACT
   Output ipValue:
   - Activation: exactly four nonempty decimal octets, each 0..255, separated by '.' (PUB001, PUB002).
   - Retention/hold: none; recomputed every scan from ipText.
   - Reset/deactivation: any malformed, nondigit, wrong-count, empty-segment, or out-of-range input yields 0 (PUB004).
   - Same-scan priority: one unconditional recomputation/write; valid 0.0.0.0 also yields 0.
   - Units/boundaries: UDINT; first octet occupies bits 31..24 and fourth bits 7..0 (PUB003).
   - Leading zeros are accepted as unspecified; each octet is limited to 3 decimal digits.
*)
FUNCTION_BLOCK FB_IPv4Parser
VAR_INPUT
    ipText : STRING(254);
END_VAR
VAR_OUTPUT
    ipValue : UDINT;
END_VAR
VAR
    strLen      : INT;
    idx         : INT;
    ch          : BYTE;
    segIndex    : INT;
    segValue    : UDINT;
    digitCount  : INT;
    accumValue  : UDINT;
END_VAR

ipValue := 0;
strLen := LEN(ipText);

IF (strLen < 7) OR (strLen > 15) THEN
    RETURN;
END_IF;

segIndex := 1;
segValue := 0;
digitCount := 0;
accumValue := 0;

FOR idx := 1 TO strLen DO
    ch := ipText[idx];

    IF (ch >= 48) AND (ch <= 57) THEN
        digitCount := digitCount + 1;
        IF digitCount > 3 THEN
            RETURN;
        END_IF;

        segValue := (segValue * 10) + (BYTE_TO_UDINT(ch) - 48);
        IF segValue > 255 THEN
            RETURN;
        END_IF;

    ELSIF ch = 46 THEN
        IF digitCount = 0 THEN
            RETURN;
        END_IF;

        IF segIndex >= 4 THEN
            RETURN;
        END_IF;

        accumValue := (accumValue * 256) + segValue;
        segIndex := segIndex + 1;
        segValue := 0;
        digitCount := 0;

    ELSE
        RETURN;
    END_IF;
END_FOR;

IF digitCount = 0 THEN
    RETURN;
END_IF;

IF segIndex <> 4 THEN
    RETURN;
END_IF;

ipValue := (accumValue * 256) + segValue;

END_FUNCTION_BLOCK

(* ---- public-medium-08.raw_candidate_01.st ---- *)
(* ENGINEERING_CONTRACT
   Output ipValue:
   - Activation: exactly four nonempty decimal octets, each 0..255, separated by '.' (PUB001, PUB002).
   - Retention/hold: none; recomputed every scan from ipText.
   - Reset/deactivation: any malformed, nondigit, wrong-count, empty-segment, or out-of-range input yields 0 (PUB004).
   - Same-scan priority: one unconditional recomputation/write; valid 0.0.0.0 also yields 0.
   - Units/boundaries: UDINT; first octet occupies bits 31..24 and fourth bits 7..0 (PUB003).
   - Leading zeros are accepted as unspecified; each octet is limited to 3 decimal digits.
*)
FUNCTION_BLOCK FB_IPv4Parser
VAR_INPUT
    ipText : STRING(254);
END_VAR
VAR_OUTPUT
    ipValue : UDINT;
END_VAR
VAR
    strLen      : INT;
    idx         : INT;
    ch          : BYTE;
    segIndex    : INT;
    segValue    : UDINT;
    digitCount  : INT;
    accumValue  : UDINT;
END_VAR

ipValue := 0;
strLen := LEN(ipText);

IF (strLen < 7) OR (strLen > 15) THEN
    RETURN;
END_IF

segIndex := 1;
segValue := 0;
digitCount := 0;
accumValue := 0;

FOR idx := 1 TO strLen DO
    ch := ipText[idx];

    IF (ch >= 48) AND (ch <= 57) THEN
        digitCount := digitCount + 1;
        IF digitCount > 3 THEN
            RETURN;
        END_IF

        segValue := (segValue * 10) + (BYTE_TO_UDINT(ch) - 48);
        IF segValue > 255 THEN
            RETURN;
        END_IF

    ELSIF ch = 46 THEN
        IF digitCount = 0 THEN
            RETURN;
        END_IF

        IF segIndex >= 4 THEN
            RETURN;
        END_IF

        accumValue := (accumValue * 256) + segValue;
        segIndex := segIndex + 1;
        segValue := 0;
        digitCount := 0;

    ELSE
        RETURN;
    END_IF
END_FOR

IF digitCount = 0 THEN
    RETURN;
END_IF

IF segIndex <> 4 THEN
    RETURN;
END_IF

ipValue := (accumValue * 256) + segValue;

END_FUNCTION_BLOCK
